(* IEC 61131-3 sources: 2026_Projet_YGO_ExcavatriceDragage/CODE_BACKUP/CODE_20260902_JoyAvantHoming_v0.6.27/G_CYCLE/_TYPES, 14 files *)

(* ---- E_CycleStep.st ---- *)
(* =======================================================================
   ⚙️ E_CycleStep — Étapes de la machine d'état du cycle automatique
   ───────────────────────────────────────────────────────────────
   🎯 Rôle : Énumération des étapes du cycle automatique de dragage (X0 à X13 + STABILIZING)
   📄 Doc métier : DOC/AF/AF_Partie-04_Mode_SemiAuto_Sequenceur_v2.3.md
   ======================================================================= *)

TYPE E_CycleStep :
(
  X0_PREPARATION      := 0,   (* Début de graphe : à la TRÉMIE, treuils en position HAUTE *)
  X1_HOMING           := 1,   (* Vitesses lentes pour chercher capteur top + référencement *)
  X2_WORK_POS_SELECT  := 2,   (* Sélection cible Trémie/P1/Maintenance + translation validée *)
  X3_OPEN_BUCKET      := 3,   (* Ouverture benne (si déjà ouverte -> passe vite) *)
  X4_DESCEND_OPEN     := 4,   (* Plongée benne ouverte, M1+M2 synchro, Kobold mesure ON *)
  X5_BOTTOM_CONFIRMED := 5,   (* Fond validé (FB_DiveSearch) ; arrêt descente *)
  X6_CLOSE_BUCKET     := 6,   (* Fermeture benne — tolérance « à peu près fermé » *)
  X7_CTRL_ASCENT      := 7,   (* Remontée palier 1 de contrôle *)
  X8_ASCENT_LOADED    := 8,   (* Remontée nominale jusqu'à limite haute *)
  X9_DRAIN_PAUSE      := 9,   (* Égouttage temporisé — temps affiché IHM *)
  X10_TRANSLATE_DUMP  := 10,  (* Translation vers trémie + avertissements IHM *)
  X11_OPEN_DUMP       := 11,  (* Ouverture benne = vidage ; montée possible, descente ouvre *)
  X13_DONE_SYNC       := 13,  (* Fin de cycle, synchronisation finale (R4) + compteur *)
  STABILIZING         := 14   (* État d'attente/stabilisation — pas une erreur *)
);
END_TYPE

(* ---- E_DiveSearchState.st ---- *)
(* =======================================================================
   ⚙️ E_DiveSearchState — Phases internes de recherche du fond Kobold
   ───────────────────────────────────────────────────────────────
   🎯 Rôle : Énumération des phases de détection et recherche du fond
   📄 Doc métier : DOC/AF/AF_Partie-04_Mode_SemiAuto_Sequenceur_v2.3.md
   ======================================================================= *)

TYPE E_DiveSearchState :
(
    WAIT_PRECONDITIONS := 0, (* Attente benne ouverte, positions et Kobold au repos *)
    READY_TO_DESCEND   := 1, (* Prêt à assister une demande de descente *)
    SEARCHING_IMMERSION := 2, (* Descending : attente front 0->1 dans fenêtre eau *)
    SEARCHING_BOTTOM    := 3, (* Immersion validée : attente front 1->0 au fond *)
    BOTTOM_CONFIRMED    := 4, (* Fond validé ; extraction peut être demandée *)
    ERROR_HOLD          := 5  (* Séquence invalide, descente assistée interdite *)
);
END_TYPE

(* ---- E_ExtractionAssistState.st ---- *)
(* =======================================================================
   ⚙️ E_ExtractionAssistState — Phases d'extraction assistée
   ───────────────────────────────────────────────────────────────
   🎯 Rôle : Énumération des phases de la séquence d'extraction assistée
   📄 Doc métier : DOC/AF/AF_Partie-04_Mode_SemiAuto_Sequenceur_v2.3.md
   ======================================================================= *)

TYPE E_ExtractionAssistState :
(
    WAIT_BOTTOM_CONFIRMATION := 0, (* Attente fond Kobold ou attestation opérateur *)
    READY_TO_CLOSE            := 1, (* Prêt à fermer la benne *)
    CLOSING_BUCKET            := 2, (* FB_Bucket ferme M2 seul *)
    CONTROL_ASCENT            := 3, (* M1/M2 synchronisés au palier sans contacteur vitesse *)
    NOMINAL_ASCENT            := 4, (* Ascending couplée avec vitesse demandée opérateur *)
    ERROR_HOLD                := 5  (* Défaut extraction, reprise interdite avant reset *)
);
END_TYPE

(* ---- E_MachineHomingStep.st ---- *)
(* =======================================================================
   ⚙️ E_MachineHomingStep — Etapes du guide de referencement machine
   ───────────────────────────────────────────────────────────────
   🎯 Rôle : Etat publie du guide de homing conjoint M1/M2/benne (IHM + interlocks)
   📄 Doc métier : DOC/AF/AF_Partie-09_Fonction_Encoder_v2.4.md (F09.08)
   ======================================================================= *)

TYPE E_MachineHomingStep :
(
    IDLE                 := 0,   (* Referencement indisponible (Enable=FALSE) *)
    LOSS_SAFESTOP        := 5,   (* Perte de datum en mouvement : arret controle en cours *)
    BOTH_NOT_HOMED       := 10,  (* Codeurs M1 et M2 non references : passer en MAINT_N2 *)
    M1_NOT_HOMED         := 11,  (* Codeur M1 non reference ou mesure douteuse : homer M1 *)
    M2_NOT_HOMED         := 12,  (* Codeur M2 non reference ou mesure douteuse : homer M2 *)
    OFFSET_UNKNOWN       := 20,  (* Offset benne inconnu : passer en MAINT_N2 *)
    NEED_TOP_POSITION    := 30,  (* Monter Both a vitesse lente jusqu au capteur haut *)
    NEED_MECHANICAL_STOP := 40,  (* Capteur haut atteint : relacher la commande et attendre l arret *)
    AWAIT_BUCKET_CONFIRM := 45,  (* Confirmer visuellement la benne : Fermee ou Ouverte *)
    HOMING_IN_PROGRESS   := 50,  (* Referencement conjoint M1/M2 en cours : ne pas manoeuvrer *)
    VALID                := 60,  (* Referencement machine valide : mode nominal disponible *)
    FAILED               := 70   (* Referencement incomplet : rester en N2 et recommencer *)
);
END_TYPE

(* ---- E_OperatorAxis.st ---- *)
(* =======================================================================
   ⚙️ E_OperatorAxis — Axe ou organe de pilotage attendu par le cycle
   ───────────────────────────────────────────────────────────────
   🎯 Rôle : Énumération de l'organe joystick/bouton attendu pour le mouvement
   📄 Doc métier : DOC/AF/AF_Partie-04_Mode_SemiAuto_Sequenceur_v2.3.md
   ======================================================================= *)

TYPE E_OperatorAxis :
(
    NONE        := 0, (* Aucun axe attendu (étape automatique ou arrêt) *)
    JOYSTICK_X  := 1, (* Axe X translation attendu *)
    JOYSTICK_Y  := 2, (* Axe Y treuils / plongée attendu *)
    BUTTON      := 3  (* Action bouton attendue (ex: validation, homing) *)
);
END_TYPE

(* ---- E_ProgramSequence.st ---- *)
(* =======================================================================
   ⚙️ E_ProgramSequence — Identifiant de la séquence programme active
   ───────────────────────────────────────────────────────────────
   🎯 Rôle : Identification de la séquence en cours d'exécution
   📄 Doc métier : DOC/AF/AF_Partie-04_Mode_SemiAuto_Sequenceur_v2.3.md
   ======================================================================= *)

TYPE E_ProgramSequence :
(
    NONE        := 0, (* Aucune séquence active *)
    MAIN_CYCLE  := 1, (* Cycle principal automatique de dragage X0..X13 *)
    DIVE_SEARCH := 2, (* Sous-séquence de plongée / recherche de fond *)
    EXTRACTION  := 3  (* Sous-séquence d'extraction et fermeture *)
);
END_TYPE

(* ---- ST_fbDiveSearch_Config.st ---- *)
(* =======================================================================
   ST_fbDiveSearch_Config - Reglages du cycle de recherche du fond
   ======================================================================= *)
TYPE ST_fbDiveSearch_Config :
STRUCT
    DiveSpeedMin_Mps       : REAL := 0.15;   // Vitesse minimale de calcul du timeout (m/s)
    TimeoutMarginFactor    : REAL := 1.5;    // Marge appliquee au temps theorique
    TimeoutMinCourse_M     : REAL := 1.0;    // Course minimale prise en compte (m)
    TimeoutMaxCourse_M     : REAL := 200.0;  // Course maximale prise en compte (m)
    SecToMs                : REAL := 1000.0; // Conversion secondes vers millisecondes
END_STRUCT
END_TYPE

(* ---- ST_fbDiveSearch_Inputs.st ---- *)
(* =======================================================================
   ST_fbDiveSearch_Inputs - Bus d'entree du cycle FB_DiveSearch
   ======================================================================= *)
TYPE ST_fbDiveSearch_Inputs :
STRUCT
    // === AUTORISATIONS & COMMANDE ===
    PowerContactorEngaged : BOOL;          // Chaine de puissance engagee
    Mode                  : E_Mode;        // Mode arbitre courant
    MotionRequestActive   : BOOL;          // Demande de mouvement couplee
    MotionDirection       : INT;           // Sens demande (-1 = descente)

    // === CAPTEURS & MESURES ===
    BucketIsOpen           : BOOL;          // Benne ouverte confirmee
    KoboldImmersed         : BOOL;          // Kobold immerge
    M1Position_M           : REAL;          // Position cable M1 (m)
    M2Position_M           : REAL;          // Position cable M2 (m)
    PositionsValid         : BOOL;          // Mesures M1/M2 valides
    CurrentSpeedStep       : INT;           // Palier reel courant (0..5)

    // === REGLAGES METIER ===
    DiveStartMin_M         : REAL;          // Position minimale avant descente (m)
    ImmersionUpper_M       : REAL;          // Borne haute fenetre immersion (m)
    ImmersionLower_M       : REAL;          // Borne basse fenetre immersion (m)
    CableLimitAscent_M     : REAL;          // Limite haute exploitation (m)
    LimitLegalDepthMin_M   : REAL;          // Limite basse legale (m)
    CfgDiveFloorStep       : INT;           // Plancher palier descente (0..5)
    CycleTime              : TIME;          // Periode d'execution du cycle
    BypassPreconditions     : BOOL;         // Bypass reserve au mode maintenance N2/test
    Config                 : ST_fbDiveSearch_Config; // Parametres timeout
END_STRUCT
END_TYPE

(* ---- ST_fbDiveSearch_Outputs.st ---- *)
(* =======================================================================
   ST_fbDiveSearch_Outputs - Bus de sortie du cycle FB_DiveSearch
   ======================================================================= *)
TYPE ST_fbDiveSearch_Outputs :
STRUCT
    // === ETAT DU CYCLE ===
    StepState              : E_DiveSearchState; // Etape courante
    StepAtFault            : E_DiveSearchState; // Etape figee au defaut

    // === PERMIS & ORDRES ASSISTES ===
    DescendPermit          : BOOL;          // Autorisation de descente assistee
    KoboldContactorCmd     : BOOL;          // Commande alimentation Kobold (fail-safe, coupe au front de fond)
    BottomTouchConfirmed   : BOOL;          // Fond confirme
    MinStepDown            : INT;           // Plancher palier descente

    // === DIAGNOSTIC OPERATEUR ===
    OperatorActionId       : WORD;          // Identifiant numerique de l'action
    OperatorAction          : STRING(120);  // Consigne operateur ASCII
END_STRUCT
END_TYPE

(* ---- ST_fbMachineHomingCycle_AxisHomingStatus.st ---- *)
(* =======================================================================
   🔌 ST_fbMachineHomingCycle_AxisHomingStatus — Statut homing d'un axe treuil
   ───────────────────────────────────────────────────────────────
   🎯 Rôle : Regroupe l'etat de homing d'un axe (M1 ou M2) consomme par
             FB_MachineHomingCycle pour piloter le guide et la transaction.
   📄 Doc métier : DOC/AF/AF_Partie-09_Fonction_Encoder_v2.4.md (F09.08)
   ======================================================================= *)
TYPE ST_fbMachineHomingCycle_AxisHomingStatus :
STRUCT
    HomedAndReliable : BOOL;   (* Codeur reference ET mesure jugee fiable (gate strict) *)
    HomingBusy       : BOOL;   (* Sequence de homing en cours sur l'axe *)
    HomingDone       : BOOL;   (* Homing termine avec succes (HomingLifecycle.Done cote FB_Encoder) *)
    HomingError      : BOOL;   (* Homing en erreur sur l'axe (HomingFault.Error) *)
END_STRUCT
END_TYPE

(* ---- ST_fbMachineHomingCycle_BucketCommit.st ---- *)
(* =======================================================================
   🔌 ST_fbMachineHomingCycle_BucketCommit — Commit atomique de l'etat benne
   ───────────────────────────────────────────────────────────────
   🎯 Rôle : Impulsion 1 scan emise par FB_MachineHomingCycle vers FB_Bucket
             apres succes des DEUX homings. FB_Bucket reste seul proprietaire
             de IsOpen / IsClosed.
   🔒 Sécurité : CommitOpen et CommitClose mutuellement exclusifs (garanti
                 par le corps du FB — rejet du double-confirm, cf. C-2).
   📄 Doc métier : DOC/AF/AF_Partie-05_Modes_Maintenance_v2.1.md
   ======================================================================= *)
TYPE ST_fbMachineHomingCycle_BucketCommit :
STRUCT
    CommitOpen  : BOOL;   (* Publier "benne ouverte" (impulsion 1 scan) *)
    CommitClose : BOOL;   (* Publier "benne fermee" (impulsion 1 scan) *)
END_STRUCT
END_TYPE

(* ---- ST_fbMachineHomingCycle_Cfg.st ---- *)
(* =======================================================================
   ⚙️ ST_fbMachineHomingCycle_Cfg — Réglages de FB_MachineHomingCycle
   ───────────────────────────────────────────────────────────────────────
   🎯 Rôle : Regrouper les réglages géométriques du référencement machine
             (cible haute M1 + écarts benne ouverte/fermée).
   🔒 Ownership : produit par le call-site PRG_02_Acquisition depuis
             _WinchM1CfgPersist et _BucketCfgPersist (GVL_PERSISTENT).
   📄 Doc : DOC/AF/AF_Partie-09_Fonction_Encoder_v2.4.md (F09.08)
   ======================================================================= *)

TYPE ST_fbMachineHomingCycle_Cfg :
STRUCT
    CfgTopHomingTarget_M : REAL;   // Cible haute configurée M1 (m)
    CfgOffsetOpen_M      : REAL;   // Ecart géométrique benne ouverte (m)
    CfgOffsetClose_M     : REAL;   // Ecart géométrique benne fermée (m)
END_STRUCT
END_TYPE

(* ---- ST_fbMachineHomingCycle_HomingDemand.st ---- *)
(* =======================================================================
   🔌 ST_fbMachineHomingCycle_HomingDemand — Demande de homing conjoint vers un axe
   ───────────────────────────────────────────────────────────────
   🎯 Rôle : Ordre de prise d'origine emis par FB_MachineHomingCycle vers
             une facade FB_Encoder. M1 : cible configuree. M2 : cible
             geometrique dynamique (top M1 configure +/- offset benne),
             jamais une position M1 live.
   📄 Doc métier : DOC/AF/AF_Partie-09_Fonction_Encoder_v2.4.md (F09.08)
   ======================================================================= *)
TYPE ST_fbMachineHomingCycle_HomingDemand :
STRUCT
    HomeReq          : BOOL;   (* Demande de prise d'origine pour cet axe (vocab reserve Homing) *)
    UseDynamicTarget : BOOL;   (* TRUE => cible = DynamicTarget_M (M2 uniquement) *)
    DynamicTarget_M  : REAL;   (* Cible geometrique benne (m) : CfgTopHomingTargetM + offset *)
END_STRUCT
END_TYPE

(* ---- ST_MachineHoming.st ---- *)
(* =======================================================================
   🧭 ST_MachineHoming — Etat publie du homing conjoint machine (M1/M2/benne)
   ───────────────────────────────────────────────────────────────
   🎯 Rôle : Regroupe les 8 sorties homing a plat de PRG_02_Acquisition en
             un bus struct unique, publie sur le bus inter-PRG.
   🔒 Sécurité : Homed = qualification conjointe reference machine (gate SEMI_AUTO).
                 HomingLoss = perte reference en mouvement : arret controle SafeStop.
   📄 Doc métier : DOC/AF/AF_Partie-09_Fonction_Encoder_v2.4.md (F09.08)
   ======================================================================= *)
TYPE ST_MachineHoming :
STRUCT
    Homed            : BOOL;          (* Qualification conjointe reference machine *)
    SetPosBucketOpen : BOOL;          (* Valider position actuelle = reference benne ouverte *)
    SetPosBucketClose: BOOL;          (* Valider position actuelle = reference benne fermee *)
    Active           : BOOL;          (* Homing conjoint en cours *)
    HomingLoss       : BOOL;          (* Perte reference en mouvement : arret controle SafeStop *)
    Step             : INT;           (* Etape guidee reference *)
    Instruction      : STRING(120);   (* Consigne IHM reference *)
    Failed           : BOOL;          (* Transaction reference abandonnee *)
END_STRUCT
END_TYPE
